// TIA Portal V21 export
// export: Created 2026-11-10T07:35:12.558758Z, ExportSetting WithDefaults, DisplayName Totally Integrated Automation Portal, DisplayVersion V21 Update 3, DisplayName STEP 7 Professional, DisplayVersion V21 Update 3, DisplayName STEP 7 Safety, DisplayVersion V21, DisplayName Tech WebApplication, DisplayVersion V21, DisplayName WinCC Basic/Comfort/Advanced, DisplayVersion V21 Update 3, DisplayName WinCC Unified, DisplayVersion V21 Update 3
FUNCTION_BLOCK "FB_Lad_ex106"   // FB31, LAD
{ S7_Optimized_Access := 'TRUE' }
VERSION : 0.1
// stored: AutoNumber true, IsIECCheckEnabled false, IsRetainMemResEnabled false, MemoryReserve 100, SetENOAutomatically false, UDAEnableTagReadback false
   VAR_INPUT
      v_ob_nr : OB_TOD;
      v_ret_val : Int;
   END_VAR
BEGIN

REGION Network 1: CAN_TINT - Cancel time-of-day interrupt
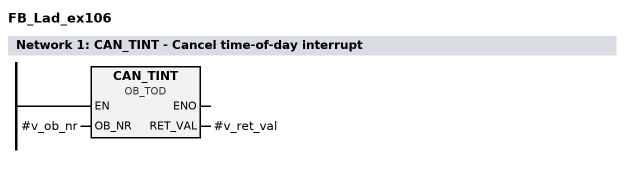
   RUNG wire#powerrail
      { S7_Templates := "ob_type := OB_TOD" } CAN_TINT(OB_NR := #v_ob_nr, Ret_Val => #v_ret_val)
   END_RUNG
   // the same network as SCL:
   #v_ret_val := CAN_TINT(OB_NR := #v_ob_nr);
END_REGION
END_FUNCTION_BLOCK
